FUNCTION_BLOCK InitState (* Basic Function Block Type *)
  (* Standard: 61499-2 *)
  (* Version 0.0, 10/21/2026, macie, Schneider Electric, Template *)
  PACKAGE Main;
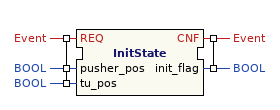
  EVENT_INPUT
    REQ WITH pusher_pos, tu_pos; (* Normal Execution Request *)
  END_EVENT
  EVENT_OUTPUT
    CNF WITH init_flag; (* Execution Confirmation *)
  END_EVENT
  VAR_INPUT
    pusher_pos : BOOL;
    tu_pos : BOOL;
  END_VAR
  VAR_OUTPUT
    init_flag : BOOL; (* Output event qualifier *)
  END_VAR
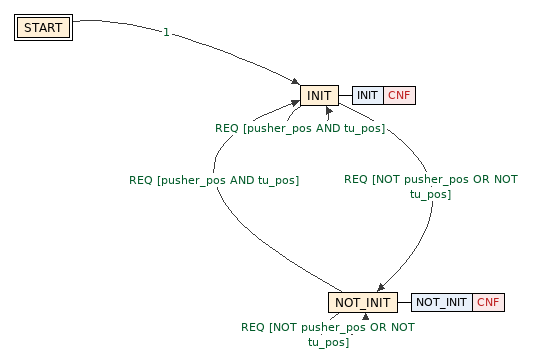
  EC_STATES
    START; (* Initial State *)
    INIT : INIT -> CNF; (* Normal execution *)
    NOT_INIT : NOT_INIT -> CNF;
  END_STATES
  EC_TRANSITIONS
    START TO INIT := 1;
    INIT TO NOT_INIT := REQ [NOT pusher_pos OR NOT tu_pos];
    NOT_INIT TO INIT := REQ [pusher_pos AND tu_pos];
    NOT_INIT TO NOT_INIT := REQ [NOT pusher_pos OR NOT tu_pos];
    INIT TO INIT := REQ [pusher_pos AND tu_pos];
  END_TRANSITIONS
  ALGORITHM INIT IN ST: (* Initialization algorithm *)
;
init_flag := TRUE;
  END_ALGORITHM
  ALGORITHM NOT_INIT IN ST: (* Normally executed algorithm *)
;
init_flag := FALSE;
  END_ALGORITHM
END_FUNCTION_BLOCK
